(* IEC 61131-3 sources: tsplc/examples/bottling-line/raw-st/src/hardware, 2 files *)

(* ---- T_Registers.st ---- *)
TYPE T_Registers : ARRAY [0..7] OF WORD;
END_TYPE

(* ---- U_Register.st ---- *)
TYPE U_Register :
UNION
	Bits : DWORD;
	Measurement : REAL;
END_UNION
END_TYPE
